(* IEC 61131-3 sources: rusty/tests/lit/multi/external_unit_linkage/interface_constructors/includer, 1 file *)

(* ---- includer.st ---- *)
FUNCTION includer : DINT
VAR_INPUT
    x : DINT;
END_VAR
    includer := x;
END_FUNCTION
